// TIA Portal V19 export
TYPE "ST_System_IO"
   STRUCT
      INPUT_BYTE : "ST_Bit";
   END_STRUCT;
END_TYPE
